(* PLC project PI_D, Desconhecido Sem nome 1 *)
(* stored: creationDateTime 2023-09-16T14:47:09, modificationDateTime 2026-11-24T21:42:17 *)

PROGRAM PI_D
  VAR
    SC : UINT;  (* OUT ANALOG PWM *)
  END_VAR
  VAR
    VP AT %IW0 : UINT;  (* INPUT ANALOG UNO A0 *)
    SP AT %QW0 : UINT;  (* SP ANALOG *)
    SO AT %QW1 : UINT := 6800;  (* SO ANALOG PWM UNO PIN10 *)
  END_VAR
  VAR
    SO_AUX : UINT;  (* SO AUXILIAR NO OUTUPUT TRACKING *)
  END_VAR
  VAR
    MF AT %QX0.0 : BOOL := 0;  (* OUT DIGITAL UNO PIN 7, MALHA FECHADA=1 *)
  END_VAR
  VAR
    VP_PERC : REAL;  (* VARIÁVEL DE PROCESSO % *)
    SP_PERC : REAL;  (* SETPOINT % *)
    SO_PERC : REAL;  (* SAÍDA DO OPERADOR % *)
    SC_PERC : REAL;  (* SAÍDA DO CONTROLADOR % *)
    SO_MAIS_P_INT_DER_PERC : REAL;  (* S0 + P+I+D % *)
    ERRO_PERC : REAL;  (* ERRO_PERC *)
    Kp_ERRO_PERC : REAL;  (* kp*ERRO_PERC *)
    Ki_ERRO_PERC : REAL;  (* kp*(1/Ti)*ERRO_PERC *)
    Ki_intgrERRO_PERC : REAL;  (* kp*(1/Ti)*intgrERRO_PERC *)
    Kd_VP_PERC : REAL;  (* kp*Td*VP_PERC *)
    Kd_derVP_PERC : REAL;  (* kp*Td*derVP_PERC *)
    M_ACAO : REAL := 1.0;  (* MODO DE AÇÃO: REVERSO=1 E DIRETO=-1 *)
    kp : REAL := 3.523;  (* BANDA PROPORCIONAL %=100/kp *)
    ki : REAL := 0.03872;  (* kp*(1/Ti) SEGUNDOS^-1 *)
    kd : REAL := 39.16;  (* kp*Td SEGUNDOS *)
    STOP_INTGR : BOOL := 0;  (* ANTI RESET WINDUP *)
    INTEGRAL_SEM_CI : INTEGRAL;
    DERIVADA : DERIVATIVE;
    SP_ant : REAL := 0.0;  (* MEMÓRIA DO SP ANTERIOR *)
    var_SP : REAL := 0.0;  (* VARIAÇÃO DO SP *)
    alfa : REAL := 1.0;  (* PARÂMETRO DO FF2GL =0 I_PD; =1 PI_D *)
    FF2GL : REAL := 0.0;  (* FEEDFORWARD 2GL *)
    MMRY : UINT := 0;  (* MEMORIA DO ALFA *)
    VP_F : REAL := 0.0;  (* VP FILTRADA (PASSA-BAIXA) PARA A DERIVADA. MALHA ABERTA: VP_F=VP_PERC *)
    kf_VP : REAL := 0.017699;  (* FILTRO DA VP: kf=Ts/(tauf+Ts)=0.02/(1.11+0.02); tauf=mu*Td=1.11 s *)
  END_VAR
  VAR  (* added by the conversion: wires and edge detectors of the diagram *)
    _SEL103_OUT : REAL;
    _NE148_OUT : BOOL;
  END_VAR

(* LD diagram, written out as Structured Text *)
(* ERRO_PERC *)
(* deadband *)
(* PROPORCIONAL *)
(* INTEGRAL *)
(* DERIVADA *)
(* 1/N,ONDE TIME CYCLE=N*[TASK0=20ms]
Exemplo: Se CYCLE=100ms ENTÃO N=5 *)
(* 1/N *)
(* N *)
(* (kp_ERRO + ki_INTEGRAL_ERRO + kd_DERIVADA_-VP) *)
SO_MAIS_P_INT_DER_PERC := Kp_ERRO_PERC + Ki_intgrERRO_PERC + Kd_derVP_PERC + SO_PERC - FF2GL;
(* PI_D se alfa=1
PI_D 2GL se 0<alfa<1
I_PD se alfa=0 *)
(* ANTI RESET WINDUP, PARAR A INTEGRAÇÃO *)
(* SATURAÇÃO DO SINAL DE CONTROLE % *)
(* DEPENDE DO COOLER O MIN *)
(* MALHA FECHADA, S0=SC,OUTPUT TRACKING
SO_AUX AJUDA NA IMPLEMENTAÇÃO
MALHA ABERTA SO_AUX=SO
MALHA FECHADA S0=SC *)
(* MALHA ABERTA, SP=VP, VP TRACKING *)
SO_AUX := SEL(MF, SO, SO_AUX);
SC_PERC := LIMIT(10.0, SO_MAIS_P_INT_DER_PERC, 100.0);
STOP_INTGR := SO_MAIS_P_INT_DER_PERC >= 100.0 OR SO_MAIS_P_INT_DER_PERC <= 10.0;
SO := SEL(MF, SO, SC);
SP := SEL(MF, VP, SP);
Ki_ERRO_PERC := ERRO_PERC * ki;
(* CONVERSOES DE REAL PARA %, VICE VERSA, DE 65535 (5V)
FILTRO DE MEDIA NA MEDIDA DE VP (???) *)
VP_PERC := UINT_TO_REAL(VP) * 0.001525;
SP_PERC := UINT_TO_REAL(SP) * 0.001525;
SO_PERC := UINT_TO_REAL(SO_AUX) * 0.001525;
SC := REAL_TO_UINT(SC_PERC * 655.35);
Kd_VP_PERC := (-1.0) * VP_F * kd * M_ACAO;
DERIVADA(RUN := TRUE, XIN := Kd_VP_PERC, CYCLE := T#500ms);
Kd_derVP_PERC := DERIVADA.XOUT * 25.0;
INTEGRAL_SEM_CI(RUN := TRUE, R1 := NOT MF, XIN := SEL(STOP_INTGR, Ki_ERRO_PERC, 0.0), X0 := 0.0, CYCLE := T#500ms);
Ki_intgrERRO_PERC := INTEGRAL_SEM_CI.XOUT * 0.04;
Kp_ERRO_PERC := ERRO_PERC * kp;
_SEL103_OUT := SEL(MF, 0.0, (SP_PERC - VP_PERC) * M_ACAO);
ERRO_PERC := SEL(ABS(_SEL103_OUT) < 0.09, _SEL103_OUT, 0.0);
(* Controlador Feedforward 2 graus de liberdade

FF2GL=kp*alfa*var_SP
var_SP= SP_PERC-SP_ant *)
_NE148_OUT := SP_PERC <> SP_ant;
var_SP := SEL(MF, 0.0, SEL(_NE148_OUT, var_SP, SP_PERC - SP_ant));
SP_ant := SEL(_NE148_OUT, SP_ant, SP_PERC);
FF2GL := SEL(MF, 0.0, SEL(_NE148_OUT AND MF, 0.0, kp * (1.0 - alfa) * var_SP) + FF2GL);
MMRY := REAL_TO_UINT(alfa * 25700.0);
(* FILTRO PASSA-BAIXA NA VP ANTES DA DERIVADA (CORRECAO DO RUIDO NO SO)
VP_F = VP_F + kf_VP*(VP_PERC - VP_F), kf_VP = Ts/(tauf+Ts) = 0.02/(1.11+0.02)
MALHA ABERTA: VP_F = VP_PERC (derivada armada, sem pulso ao fechar a malha) *)
VP_F := SEL(MF, VP_PERC, VP_F + (VP_PERC - VP_F) * kf_VP);
END_PROGRAM

CONFIGURATION Config0
  RESOURCE Res0 ON PLC
    TASK task0(INTERVAL := T#20ms, PRIORITY := 0);
    PROGRAM instance0 WITH task0 : PI_D;
  END_RESOURCE
END_CONFIGURATION
